// TIA Portal V17 program export: 0 tag tables, 0 data types, 5 data blocks, 5 code blocks (in call order from the OBs), 4 instance data blocks

DATA_BLOCK "DB_HMI"   // DB1
{ S7_Optimized_Access := 'TRUE' }
VERSION : 0.1
// stored: AutoNumber true, DBAccessibleFromOPCUA true, IsOnlyStoredInLoadMemory false, IsRetainMemResEnabled false, IsWriteProtectedInAS false, MemoryReserve 100
   VAR
      Cmd_Marcha : Bool;   // Boton MARCHA de la HMI (momentaneo)
      Cmd_Paro : Bool;   // Boton PARO de la HMI (momentaneo)
      Cmd_Reset : Bool;   // Boton RESET de la HMI (momentaneo)
      Sel_Estilo : Int := 1;   // 1 Banderas, 2 Moore, 3 Mealy
      Estado : Int;   // Estado del estilo seleccionado: 0 Reposo, 10 Marcha, 90 Falla
      Motor_En_Marcha : Bool;   // Copia de KM1_Motor para la HMI
      Falla_Termico : Bool;   // Termico disparado
      Pantalla : Int;   // Pantalla activa en la HMI (1 Principal, 2 Diagnostico, 3 Estilos)
   END_VAR
BEGIN
END_DATA_BLOCK

DATA_BLOCK "DB_Mando"
{ S7_Optimized_Access := 'TRUE' }
VERSION : 0.1
NON_RETAIN
"FB_Mando_Motor"

BEGIN

END_DATA_BLOCK

DATA_BLOCK "DB_Motor_Banderas"
{ S7_Optimized_Access := 'TRUE' }
VERSION : 0.1
NON_RETAIN
"FB_Motor_Banderas"

BEGIN

END_DATA_BLOCK

DATA_BLOCK "DB_Motor_Mealy"
{ S7_Optimized_Access := 'TRUE' }
VERSION : 0.1
NON_RETAIN
"FB_Motor_Mealy"

BEGIN

END_DATA_BLOCK

DATA_BLOCK "DB_Motor_Moore"
{ S7_Optimized_Access := 'TRUE' }
VERSION : 0.1
NON_RETAIN
"FB_Motor_Moore"

BEGIN

END_DATA_BLOCK

ORGANIZATION_BLOCK "Main"   // OB1, LAD, ProgramCycle
TITLE = "Main Program Sweep (Cycle)" / Programa principal - Arranque y paro v2
{ S7_Optimized_Access := 'TRUE' }
VERSION : 0.1
// OB1 director: una red por función. Los 3 estilos corren a la vez; el selector de la HMI decide cuál maneja KM1 y los pilotos.
// stored: AutoNumber true, IsIECCheckEnabled false, SetENOAutomatically false
   VAR_INPUT
      Initial_Call : Bool;   // Initial call of this OB
      Remanence : Bool;   // =True, if remanent data are available
   END_VAR
BEGIN

REGION Network 1: MANDO: pulsadores + HMI
   // Une entradas físicas y botones de la HMI.
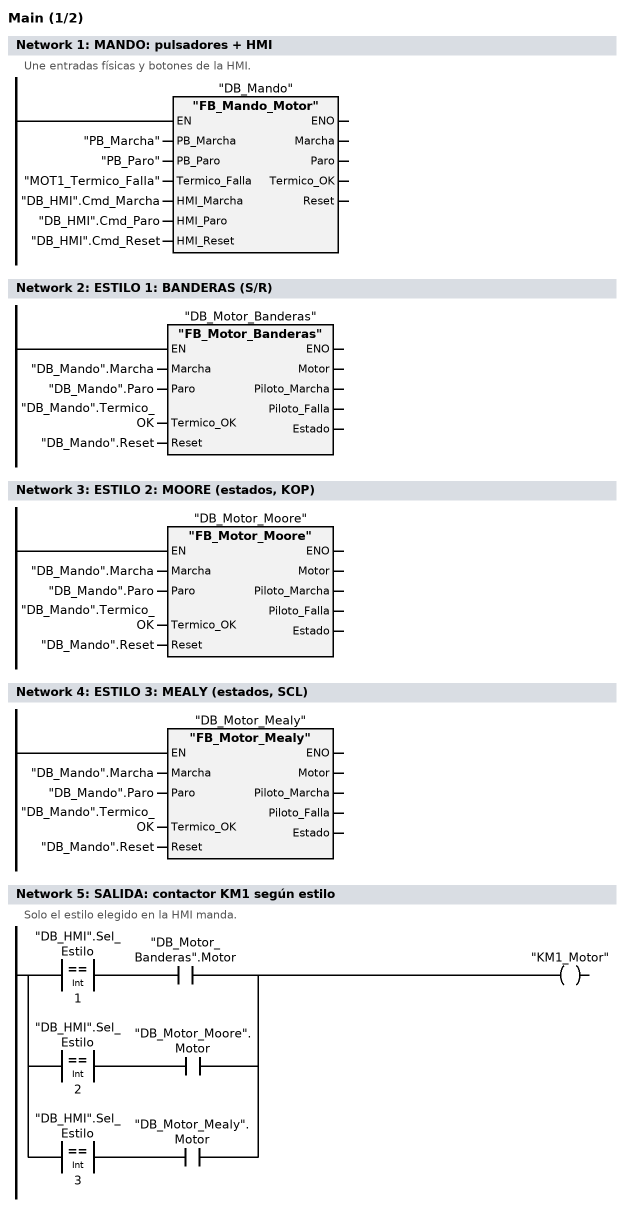
   RUNG wire#powerrail
      "DB_Mando"(PB_Marcha := "PB_Marcha", PB_Paro := "PB_Paro", Termico_Falla := "MOT1_Termico_Falla", HMI_Marcha := "DB_HMI".Cmd_Marcha, HMI_Paro := "DB_HMI".Cmd_Paro, HMI_Reset := "DB_HMI".Cmd_Reset, Marcha =>, Paro =>, Termico_OK =>, Reset =>)
   END_RUNG
   // the same network as SCL:
   "DB_Mando"(PB_Marcha := "PB_Marcha",   // "FB_Mando_Motor"
              PB_Paro := "PB_Paro",
              Termico_Falla := "MOT1_Termico_Falla",
              HMI_Marcha := "DB_HMI".Cmd_Marcha,
              HMI_Paro := "DB_HMI".Cmd_Paro,
              HMI_Reset := "DB_HMI".Cmd_Reset);
END_REGION

REGION Network 2: ESTILO 1: BANDERAS (S/R)
   RUNG wire#powerrail
      "DB_Motor_Banderas"(Marcha := "DB_Mando".Marcha, Paro := "DB_Mando".Paro, Termico_OK := "DB_Mando".Termico_OK, Reset := "DB_Mando".Reset, Motor =>, Piloto_Marcha =>, Piloto_Falla =>, Estado =>)
   END_RUNG
   // the same network as SCL:
   "DB_Motor_Banderas"(Marcha := "DB_Mando".Marcha,   // "FB_Motor_Banderas"
                       Paro := "DB_Mando".Paro,
                       Termico_OK := "DB_Mando".Termico_OK,
                       Reset := "DB_Mando".Reset);
END_REGION

REGION Network 3: ESTILO 2: MOORE (estados, KOP)
   RUNG wire#powerrail
      "DB_Motor_Moore"(Marcha := "DB_Mando".Marcha, Paro := "DB_Mando".Paro, Termico_OK := "DB_Mando".Termico_OK, Reset := "DB_Mando".Reset, Motor =>, Piloto_Marcha =>, Piloto_Falla =>, Estado =>)
   END_RUNG
   // the same network as SCL:
   "DB_Motor_Moore"(Marcha := "DB_Mando".Marcha,   // "FB_Motor_Moore"
                    Paro := "DB_Mando".Paro,
                    Termico_OK := "DB_Mando".Termico_OK,
                    Reset := "DB_Mando".Reset);
END_REGION

REGION Network 4: ESTILO 3: MEALY (estados, SCL)
   RUNG wire#powerrail
      "DB_Motor_Mealy"(Marcha := "DB_Mando".Marcha, Paro := "DB_Mando".Paro, Termico_OK := "DB_Mando".Termico_OK, Reset := "DB_Mando".Reset, Motor =>, Piloto_Marcha =>, Piloto_Falla =>, Estado =>)
   END_RUNG
   // the same network as SCL:
   "DB_Motor_Mealy"(Marcha := "DB_Mando".Marcha,   // "FB_Motor_Mealy"
                    Paro := "DB_Mando".Paro,
                    Termico_OK := "DB_Mando".Termico_OK,
                    Reset := "DB_Mando".Reset);
END_REGION

REGION Network 5: SALIDA: contactor KM1 según estilo
   // Solo el estilo elegido en la HMI manda.
   RUNG wire#powerrail
      { S7_Templates := "SrcType := Int" } EQ_Contact(in1 := "DB_HMI".Sel_Estilo, in2 := 1)
      Contact( "DB_Motor_Banderas".Motor )
      wire#w1
      Coil( "KM1_Motor" )
   END_RUNG
   RUNG wire#powerrail
      { S7_Templates := "SrcType := Int" } EQ_Contact(in1 := "DB_HMI".Sel_Estilo, in2 := 2)
      Contact( "DB_Motor_Moore".Motor )
   END_RUNG wire#w1
   RUNG wire#powerrail
      { S7_Templates := "SrcType := Int" } EQ_Contact(in1 := "DB_HMI".Sel_Estilo, in2 := 3)
      Contact( "DB_Motor_Mealy".Motor )
   END_RUNG wire#w1
   // the same network as SCL:
   "KM1_Motor" := (("DB_HMI".Sel_Estilo = 1) AND "DB_Motor_Banderas".Motor) OR (("DB_HMI".Sel_Estilo = 2) AND "DB_Motor_Moore".Motor) OR (("DB_HMI".Sel_Estilo = 3) AND "DB_Motor_Mealy".Motor);
END_REGION

REGION Network 6: SALIDA: piloto de marcha
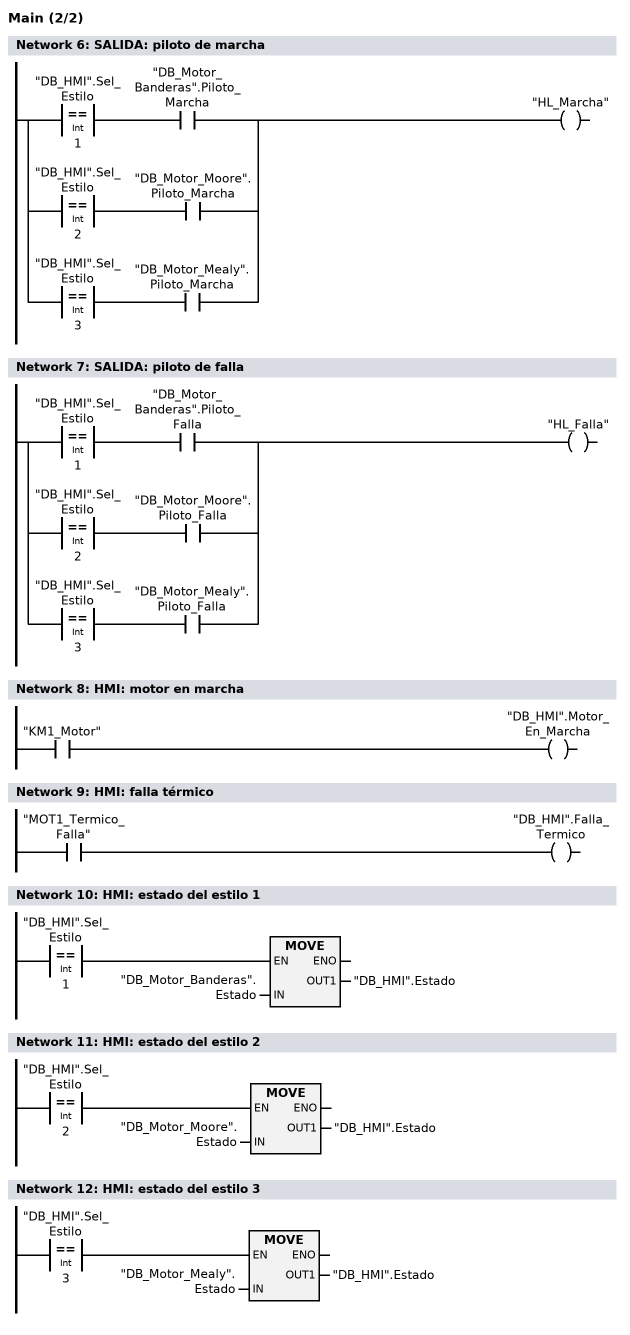
   RUNG wire#powerrail
      { S7_Templates := "SrcType := Int" } EQ_Contact(in1 := "DB_HMI".Sel_Estilo, in2 := 1)
      Contact( "DB_Motor_Banderas".Piloto_Marcha )
      wire#w1
      Coil( "HL_Marcha" )
   END_RUNG
   RUNG wire#powerrail
      { S7_Templates := "SrcType := Int" } EQ_Contact(in1 := "DB_HMI".Sel_Estilo, in2 := 2)
      Contact( "DB_Motor_Moore".Piloto_Marcha )
   END_RUNG wire#w1
   RUNG wire#powerrail
      { S7_Templates := "SrcType := Int" } EQ_Contact(in1 := "DB_HMI".Sel_Estilo, in2 := 3)
      Contact( "DB_Motor_Mealy".Piloto_Marcha )
   END_RUNG wire#w1
   // the same network as SCL:
   "HL_Marcha" := (("DB_HMI".Sel_Estilo = 1) AND "DB_Motor_Banderas".Piloto_Marcha) OR (("DB_HMI".Sel_Estilo = 2) AND "DB_Motor_Moore".Piloto_Marcha) OR (("DB_HMI".Sel_Estilo = 3) AND "DB_Motor_Mealy".Piloto_Marcha);
END_REGION

REGION Network 7: SALIDA: piloto de falla
   RUNG wire#powerrail
      { S7_Templates := "SrcType := Int" } EQ_Contact(in1 := "DB_HMI".Sel_Estilo, in2 := 1)
      Contact( "DB_Motor_Banderas".Piloto_Falla )
      wire#w1
      Coil( "HL_Falla" )
   END_RUNG
   RUNG wire#powerrail
      { S7_Templates := "SrcType := Int" } EQ_Contact(in1 := "DB_HMI".Sel_Estilo, in2 := 2)
      Contact( "DB_Motor_Moore".Piloto_Falla )
   END_RUNG wire#w1
   RUNG wire#powerrail
      { S7_Templates := "SrcType := Int" } EQ_Contact(in1 := "DB_HMI".Sel_Estilo, in2 := 3)
      Contact( "DB_Motor_Mealy".Piloto_Falla )
   END_RUNG wire#w1
   // the same network as SCL:
   "HL_Falla" := (("DB_HMI".Sel_Estilo = 1) AND "DB_Motor_Banderas".Piloto_Falla) OR (("DB_HMI".Sel_Estilo = 2) AND "DB_Motor_Moore".Piloto_Falla) OR (("DB_HMI".Sel_Estilo = 3) AND "DB_Motor_Mealy".Piloto_Falla);
END_REGION

REGION Network 8: HMI: motor en marcha
   RUNG wire#powerrail
      Contact( "KM1_Motor" )
      Coil( "DB_HMI".Motor_En_Marcha )
   END_RUNG
   // the same network as SCL:
   "DB_HMI".Motor_En_Marcha := "KM1_Motor";
END_REGION

REGION Network 9: HMI: falla térmico
   RUNG wire#powerrail
      Contact( "MOT1_Termico_Falla" )
      Coil( "DB_HMI".Falla_Termico )
   END_RUNG
   // the same network as SCL:
   "DB_HMI".Falla_Termico := "MOT1_Termico_Falla";
END_REGION

REGION Network 10: HMI: estado del estilo 1
   RUNG wire#powerrail
      { S7_Templates := "SrcType := Int" } EQ_Contact(in1 := "DB_HMI".Sel_Estilo, in2 := 1)
      { S7_GenerateENO := "TRUE" } Move(in := "DB_Motor_Banderas".Estado, out1 => "DB_HMI".Estado)
   END_RUNG
   // the same network as SCL:
   IF "DB_HMI".Sel_Estilo = 1 THEN "DB_HMI".Estado := "DB_Motor_Banderas".Estado; END_IF;
END_REGION

REGION Network 11: HMI: estado del estilo 2
   RUNG wire#powerrail
      { S7_Templates := "SrcType := Int" } EQ_Contact(in1 := "DB_HMI".Sel_Estilo, in2 := 2)
      { S7_GenerateENO := "TRUE" } Move(in := "DB_Motor_Moore".Estado, out1 => "DB_HMI".Estado)
   END_RUNG
   // the same network as SCL:
   IF "DB_HMI".Sel_Estilo = 2 THEN "DB_HMI".Estado := "DB_Motor_Moore".Estado; END_IF;
END_REGION

REGION Network 12: HMI: estado del estilo 3
   RUNG wire#powerrail
      { S7_Templates := "SrcType := Int" } EQ_Contact(in1 := "DB_HMI".Sel_Estilo, in2 := 3)
      { S7_GenerateENO := "TRUE" } Move(in := "DB_Motor_Mealy".Estado, out1 => "DB_HMI".Estado)
   END_RUNG
   // the same network as SCL:
   IF "DB_HMI".Sel_Estilo = 3 THEN "DB_HMI".Estado := "DB_Motor_Mealy".Estado; END_IF;
END_REGION
END_ORGANIZATION_BLOCK

FUNCTION_BLOCK "FB_Mando_Motor"   // FB1, LAD
TITLE = Mando del motor: pulsadores + HMI
{ S7_Optimized_Access := 'TRUE' }
VERSION : 0.1
// Une pulsadores físicos y botones HMI. Reset = botón RESET de la HMI o mantener MARCHA 3 s.
// stored: AutoNumber true, IsIECCheckEnabled false, IsRetainMemResEnabled false, MemoryReserve 100, SetENOAutomatically false, UDAEnableTagReadback false
   VAR_INPUT
      PB_Marcha : Bool;   // Pulsador MARCHA (NA)
      PB_Paro : Bool;   // Pulsador PARO: 1 = pulsado
      Termico_Falla : Bool;   // Relé térmico: 1 = disparado
      HMI_Marcha : Bool;
      HMI_Paro : Bool;
      HMI_Reset : Bool;
   END_VAR
   VAR_OUTPUT
      Marcha : Bool;
      Paro : Bool;
      Termico_OK : Bool;
      Reset : Bool;
   END_VAR
   VAR
      T_Reset : TON_TIME;   // Tiempo de MARCHA mantenida
      Reset_Mantenido : Bool;   // MARCHA mantenida 3 s
   END_VAR
BEGIN

REGION Network 1: Marcha
   // Pulsador físico o botón de la HMI.
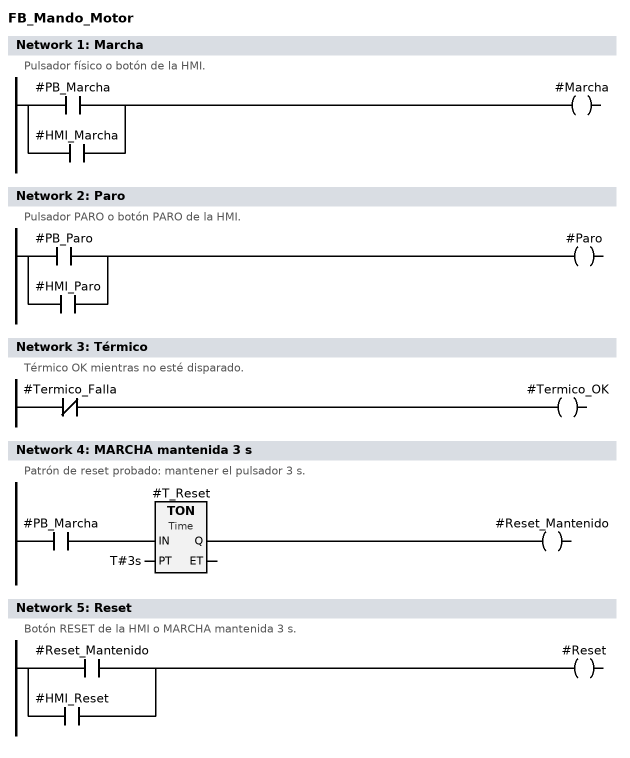
   RUNG wire#powerrail
      Contact( #PB_Marcha )
      wire#w1
      Coil( #Marcha )
   END_RUNG
   RUNG wire#powerrail
      Contact( #HMI_Marcha )
   END_RUNG wire#w1
   // the same network as SCL:
   #Marcha := #PB_Marcha OR #HMI_Marcha;
END_REGION

REGION Network 2: Paro
   // Pulsador PARO o botón PARO de la HMI.
   RUNG wire#powerrail
      Contact( #PB_Paro )
      wire#w1
      Coil( #Paro )
   END_RUNG
   RUNG wire#powerrail
      Contact( #HMI_Paro )
   END_RUNG wire#w1
   // the same network as SCL:
   #Paro := #PB_Paro OR #HMI_Paro;
END_REGION

REGION Network 3: Térmico
   // Térmico OK mientras no esté disparado.
   RUNG wire#powerrail
      I_Contact( #Termico_Falla )
      Coil( #Termico_OK )
   END_RUNG
   // the same network as SCL:
   #Termico_OK := NOT #Termico_Falla;
END_REGION

REGION Network 4: MARCHA mantenida 3 s
   // Patrón de reset probado: mantener el pulsador 3 s.
   RUNG wire#powerrail
      Contact( #PB_Marcha )
      { S7_Templates := "time_type := Time" } #T_Reset.TON(pt := T#3s, et =>)
      Coil( #Reset_Mantenido )
   END_RUNG
   // the same network as SCL:
   #T_Reset(IN := #PB_Marcha, PT := T#3s);   // TON
   #Reset_Mantenido := #T_Reset.Q;
END_REGION

REGION Network 5: Reset
   // Botón RESET de la HMI o MARCHA mantenida 3 s.
   RUNG wire#powerrail
      Contact( #Reset_Mantenido )
      wire#w1
      Coil( #Reset )
   END_RUNG
   RUNG wire#powerrail
      Contact( #HMI_Reset )
   END_RUNG wire#w1
   // the same network as SCL:
   #Reset := #Reset_Mantenido OR #HMI_Reset;
END_REGION
END_FUNCTION_BLOCK

FUNCTION_BLOCK "FB_Motor_Banderas"   // FB3, LAD
TITLE = Arranque y paro por BANDERAS (S/R)
{ S7_Optimized_Access := 'TRUE' }
VERSION : 0.1
// Estilo clásico: bandera de marcha con SET/RESET (paro dominante). Sin térmico se para; al recuperarse el térmico se puede volver a arrancar sin RESET.
// stored: AutoNumber true, IsIECCheckEnabled false, IsRetainMemResEnabled false, MemoryReserve 100, SetENOAutomatically false, UDAEnableTagReadback false
   VAR_INPUT
      Marcha : Bool;   // Orden de marcha (pulsador o HMI)
      Paro : Bool;   // Orden de paro: 1 = parar
      Termico_OK : Bool;   // 1 = relé térmico sin falla
      Reset : Bool;   // Reset de falla
   END_VAR
   VAR_OUTPUT
      Motor : Bool;   // Orden al contactor
      Piloto_Marcha : Bool;   // Piloto verde
      Piloto_Falla : Bool;   // Piloto rojo
      Estado : Int;   // 0 Reposo, 10 Marcha, 90 Falla
   END_VAR
   VAR
      B_Marcha : Bool;   // Bandera: motor en marcha
      B_Falla : Bool;   // Bandera: falla térmico
   END_VAR
BEGIN

REGION Network 1: SET bandera de marcha
   // Marcha sin paro y con térmico OK.
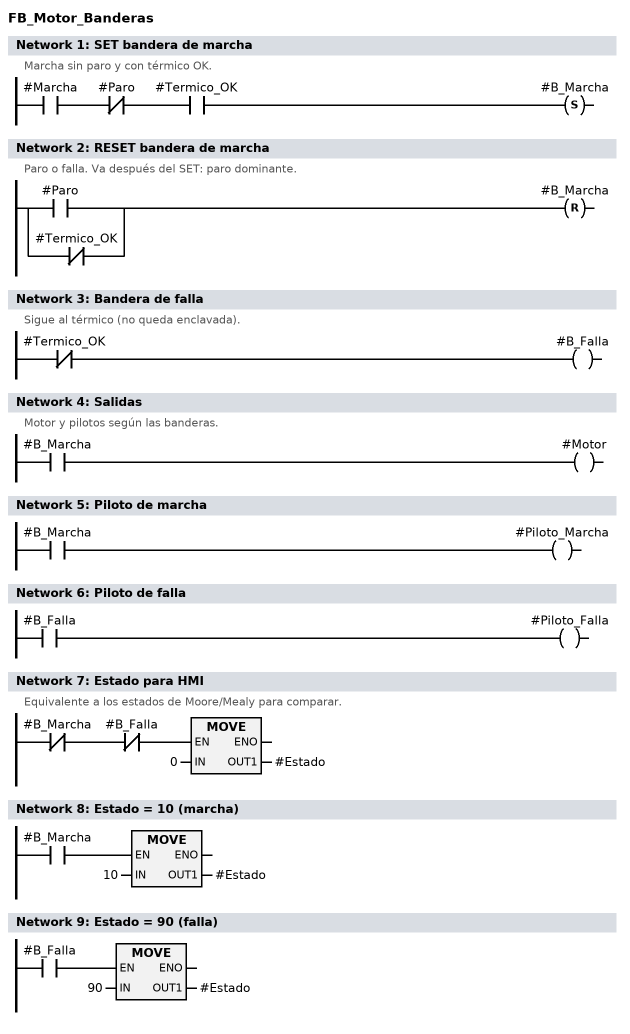
   RUNG wire#powerrail
      Contact( #Marcha )
      I_Contact( #Paro )
      Contact( #Termico_OK )
      S_Coil( #B_Marcha )
   END_RUNG
   // the same network as SCL:
   IF #Marcha AND NOT #Paro AND #Termico_OK THEN #B_Marcha := TRUE; END_IF;
END_REGION

REGION Network 2: RESET bandera de marcha
   // Paro o falla. Va después del SET: paro dominante.
   RUNG wire#powerrail
      Contact( #Paro )
      wire#w1
      R_Coil( #B_Marcha )
   END_RUNG
   RUNG wire#powerrail
      I_Contact( #Termico_OK )
   END_RUNG wire#w1
   // the same network as SCL:
   IF #Paro OR NOT #Termico_OK THEN #B_Marcha := FALSE; END_IF;
END_REGION

REGION Network 3: Bandera de falla
   // Sigue al térmico (no queda enclavada).
   RUNG wire#powerrail
      I_Contact( #Termico_OK )
      Coil( #B_Falla )
   END_RUNG
   // the same network as SCL:
   #B_Falla := NOT #Termico_OK;
END_REGION

REGION Network 4: Salidas
   // Motor y pilotos según las banderas.
   RUNG wire#powerrail
      Contact( #B_Marcha )
      Coil( #Motor )
   END_RUNG
   // the same network as SCL:
   #Motor := #B_Marcha;
END_REGION

REGION Network 5: Piloto de marcha
   RUNG wire#powerrail
      Contact( #B_Marcha )
      Coil( #Piloto_Marcha )
   END_RUNG
   // the same network as SCL:
   #Piloto_Marcha := #B_Marcha;
END_REGION

REGION Network 6: Piloto de falla
   RUNG wire#powerrail
      Contact( #B_Falla )
      Coil( #Piloto_Falla )
   END_RUNG
   // the same network as SCL:
   #Piloto_Falla := #B_Falla;
END_REGION

REGION Network 7: Estado para HMI
   // Equivalente a los estados de Moore/Mealy para comparar.
   RUNG wire#powerrail
      I_Contact( #B_Marcha )
      I_Contact( #B_Falla )
      { S7_GenerateENO := "TRUE" } Move(in := 0, out1 => #Estado)
   END_RUNG
   // the same network as SCL:
   IF NOT #B_Marcha AND NOT #B_Falla THEN #Estado := 0; END_IF;
END_REGION

REGION Network 8: Estado = 10 (marcha)
   RUNG wire#powerrail
      Contact( #B_Marcha )
      { S7_GenerateENO := "TRUE" } Move(in := 10, out1 => #Estado)
   END_RUNG
   // the same network as SCL:
   IF #B_Marcha THEN #Estado := 10; END_IF;
END_REGION

REGION Network 9: Estado = 90 (falla)
   RUNG wire#powerrail
      Contact( #B_Falla )
      { S7_GenerateENO := "TRUE" } Move(in := 90, out1 => #Estado)
   END_RUNG
   // the same network as SCL:
   IF #B_Falla THEN #Estado := 90; END_IF;
END_REGION
END_FUNCTION_BLOCK

FUNCTION_BLOCK "FB_Motor_Moore"   // FB5, LAD
TITLE = Arranque y paro: máquina de estados MOORE
{ S7_Optimized_Access := 'TRUE' }
VERSION : 0.1
// Moore: las salidas dependen solo del estado. Generado por TIA_MCP_V17 (crear_maquina_estados).
// stored: AutoNumber true, IsIECCheckEnabled false, IsRetainMemResEnabled false, MemoryReserve 100, SetENOAutomatically false, UDAEnableTagReadback false
   VAR_INPUT
      Marcha : Bool;   // Orden de marcha (pulsador o HMI)
      Paro : Bool;   // Orden de paro: 1 = parar
      Termico_OK : Bool;   // 1 = relé térmico sin falla
      Reset : Bool;   // Reset de falla
   END_VAR
   VAR_OUTPUT
      Motor : Bool;   // Orden al contactor
      Piloto_Marcha : Bool;   // Piloto verde
      Piloto_Falla : Bool;   // Piloto rojo
      Estado : Int;   // Estado actual
   END_VAR
   VAR
      Estado_Actual : Int := 0;   // Estado de la máquina
   END_VAR
   VAR_TEMP
      Estado_Previo : Int;   // Estado al inicio del ciclo
   END_VAR
BEGIN

REGION Network 1: Foto del estado al inicio del ciclo
   // Las transiciones se evalúan sobre esta copia: un solo salto por ciclo.
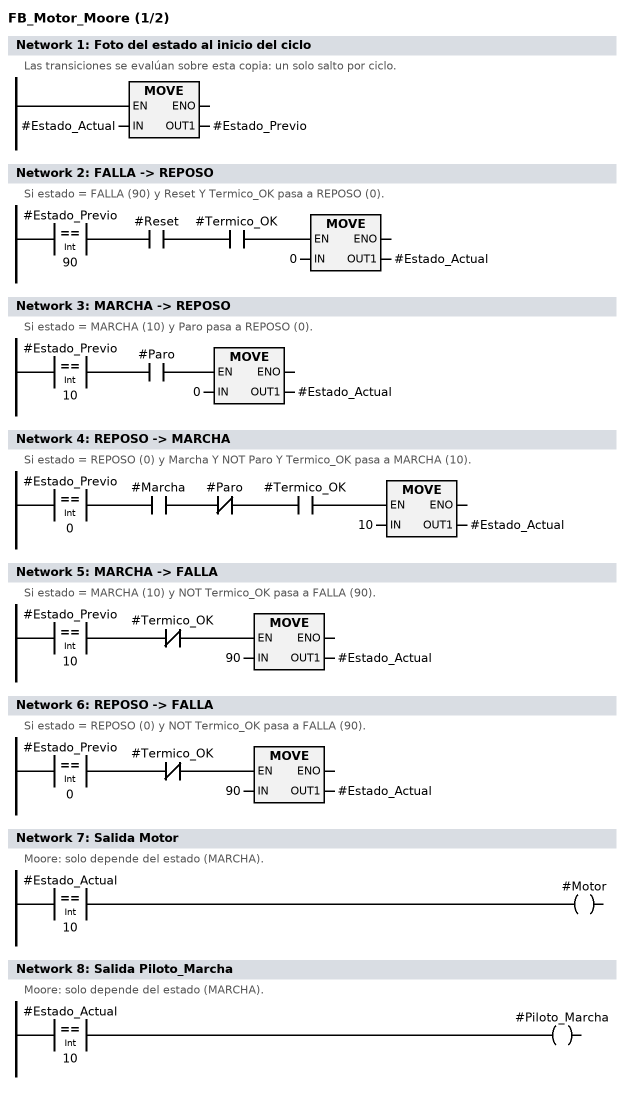
   RUNG wire#powerrail
      { S7_GenerateENO := "TRUE" } Move(in := #Estado_Actual, out1 => #Estado_Previo)
   END_RUNG
   // the same network as SCL:
   #Estado_Previo := #Estado_Actual;
END_REGION

REGION Network 2: FALLA -> REPOSO
   // Si estado = FALLA (90) y Reset Y Termico_OK pasa a REPOSO (0).
   RUNG wire#powerrail
      { S7_Templates := "SrcType := Int" } EQ_Contact(in1 := #Estado_Previo, in2 := 90)
      Contact( #Reset )
      Contact( #Termico_OK )
      { S7_GenerateENO := "TRUE" } Move(in := 0, out1 => #Estado_Actual)
   END_RUNG
   // the same network as SCL:
   IF (#Estado_Previo = 90) AND #Reset AND #Termico_OK THEN #Estado_Actual := 0; END_IF;
END_REGION

REGION Network 3: MARCHA -> REPOSO
   // Si estado = MARCHA (10) y Paro pasa a REPOSO (0).
   RUNG wire#powerrail
      { S7_Templates := "SrcType := Int" } EQ_Contact(in1 := #Estado_Previo, in2 := 10)
      Contact( #Paro )
      { S7_GenerateENO := "TRUE" } Move(in := 0, out1 => #Estado_Actual)
   END_RUNG
   // the same network as SCL:
   IF (#Estado_Previo = 10) AND #Paro THEN #Estado_Actual := 0; END_IF;
END_REGION

REGION Network 4: REPOSO -> MARCHA
   // Si estado = REPOSO (0) y Marcha Y NOT Paro Y Termico_OK pasa a MARCHA (10).
   RUNG wire#powerrail
      { S7_Templates := "SrcType := Int" } EQ_Contact(in1 := #Estado_Previo, in2 := 0)
      Contact( #Marcha )
      I_Contact( #Paro )
      Contact( #Termico_OK )
      { S7_GenerateENO := "TRUE" } Move(in := 10, out1 => #Estado_Actual)
   END_RUNG
   // the same network as SCL:
   IF (#Estado_Previo = 0) AND #Marcha AND NOT #Paro AND #Termico_OK THEN #Estado_Actual := 10; END_IF;
END_REGION

REGION Network 5: MARCHA -> FALLA
   // Si estado = MARCHA (10) y NOT Termico_OK pasa a FALLA (90).
   RUNG wire#powerrail
      { S7_Templates := "SrcType := Int" } EQ_Contact(in1 := #Estado_Previo, in2 := 10)
      I_Contact( #Termico_OK )
      { S7_GenerateENO := "TRUE" } Move(in := 90, out1 => #Estado_Actual)
   END_RUNG
   // the same network as SCL:
   IF (#Estado_Previo = 10) AND NOT #Termico_OK THEN #Estado_Actual := 90; END_IF;
END_REGION

REGION Network 6: REPOSO -> FALLA
   // Si estado = REPOSO (0) y NOT Termico_OK pasa a FALLA (90).
   RUNG wire#powerrail
      { S7_Templates := "SrcType := Int" } EQ_Contact(in1 := #Estado_Previo, in2 := 0)
      I_Contact( #Termico_OK )
      { S7_GenerateENO := "TRUE" } Move(in := 90, out1 => #Estado_Actual)
   END_RUNG
   // the same network as SCL:
   IF (#Estado_Previo = 0) AND NOT #Termico_OK THEN #Estado_Actual := 90; END_IF;
END_REGION

REGION Network 7: Salida Motor
   // Moore: solo depende del estado (MARCHA).
   RUNG wire#powerrail
      { S7_Templates := "SrcType := Int" } EQ_Contact(in1 := #Estado_Actual, in2 := 10)
      Coil( #Motor )
   END_RUNG
   // the same network as SCL:
   #Motor := #Estado_Actual = 10;
END_REGION

REGION Network 8: Salida Piloto_Marcha
   // Moore: solo depende del estado (MARCHA).
   RUNG wire#powerrail
      { S7_Templates := "SrcType := Int" } EQ_Contact(in1 := #Estado_Actual, in2 := 10)
      Coil( #Piloto_Marcha )
   END_RUNG
   // the same network as SCL:
   #Piloto_Marcha := #Estado_Actual = 10;
END_REGION

REGION Network 9: Salida Piloto_Falla
   // Moore: solo depende del estado (FALLA).
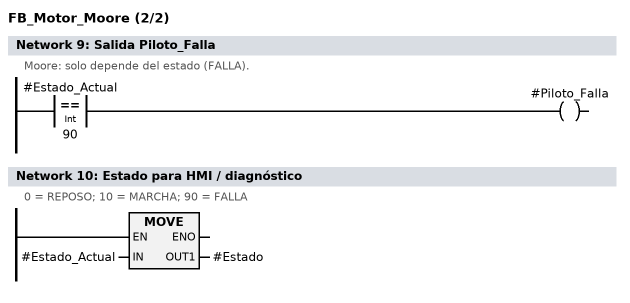
   RUNG wire#powerrail
      { S7_Templates := "SrcType := Int" } EQ_Contact(in1 := #Estado_Actual, in2 := 90)
      Coil( #Piloto_Falla )
   END_RUNG
   // the same network as SCL:
   #Piloto_Falla := #Estado_Actual = 90;
END_REGION

REGION Network 10: Estado para HMI / diagnóstico
   // 0 = REPOSO; 10 = MARCHA; 90 = FALLA
   RUNG wire#powerrail
      { S7_GenerateENO := "TRUE" } Move(in := #Estado_Actual, out1 => #Estado)
   END_RUNG
   // the same network as SCL:
   #Estado := #Estado_Actual;
END_REGION
END_FUNCTION_BLOCK

FUNCTION_BLOCK "FB_Motor_Mealy"   // FB4, SCL
TITLE = Arranque y paro: maquina de estados MEALY
{ S7_Optimized_Access := 'TRUE' }
VERSION : 0.1
// stored: AutoNumber true, IsIECCheckEnabled false, IsRetainMemResEnabled false, MemoryReserve 100, SetENOAutomatically false, UDAEnableTagReadback false
   VAR_INPUT
      Marcha : Bool;   // Orden de marcha (pulsador o HMI)
      Paro : Bool;   // Orden de paro: 1 = parar
      Termico_OK : Bool;   // 1 = rele termico sin falla
      Reset : Bool;   // Reset de falla
   END_VAR
   VAR_OUTPUT
      Motor : Bool;   // Orden al contactor
      Piloto_Marcha : Bool;   // Piloto verde
      Piloto_Falla : Bool;   // Piloto rojo
      Estado : Int;   // Estado actual (HMI)
   END_VAR
   VAR
      Estado_Actual : Int := 0;   // Estado de la maquina
   END_VAR
   VAR_TEMP
      Estado_Previo : Int;   // Estado al inicio del ciclo
   END_VAR
BEGIN
       // Mealy: las salidas dependen del estado y de las entradas (reaccion en el mismo ciclo). Generado por TIA_MCP_V17 (crear_maquina_estados).
       // Estados: 0 = REPOSO, 10 = MARCHA, 90 = FALLA

       // --- Salidas (estado actual + entradas) ---
       #Motor := (#Estado_Actual = 10 AND NOT #Paro AND #Termico_OK);
       #Piloto_Marcha := #Estado_Actual = 10;
       #Piloto_Falla := #Estado_Actual = 90;

       // --- Transiciones (sobre la foto del estado: un salto por ciclo) ---
       #Estado_Previo := #Estado_Actual;
       CASE #Estado_Previo OF
           0: // REPOSO
               IF NOT #Termico_OK THEN
                   #Estado_Actual := 90;   // -> FALLA
               ELSIF #Marcha AND NOT #Paro AND #Termico_OK THEN
                   #Estado_Actual := 10;   // -> MARCHA
               END_IF;
           10: // MARCHA
               IF NOT #Termico_OK THEN
                   #Estado_Actual := 90;   // -> FALLA
               ELSIF #Paro THEN
                   #Estado_Actual := 0;   // -> REPOSO
               END_IF;
           90: // FALLA
               IF #Reset AND #Termico_OK THEN
                   #Estado_Actual := 0;   // -> REPOSO
               END_IF;
           ELSE  // estado desconocido: volver al inicial
               #Estado_Actual := 0;
       END_CASE;

       #Estado := #Estado_Actual;
END_FUNCTION_BLOCK

DATA_BLOCK "DB_Mando"   // DB2
VERSION : 0.1
// stored: AutoNumber true, DBAccessibleFromOPCUA true, InstanceOfName FB_Mando_Motor, InstanceOfType FB
"FB_Mando_Motor"
BEGIN
END_DATA_BLOCK

DATA_BLOCK "DB_Motor_Banderas"   // DB3
VERSION : 0.1
// stored: AutoNumber true, DBAccessibleFromOPCUA true, InstanceOfName FB_Motor_Banderas, InstanceOfType FB
"FB_Motor_Banderas"
BEGIN
END_DATA_BLOCK

DATA_BLOCK "DB_Motor_Mealy"   // DB5
VERSION : 0.1
// stored: AutoNumber true, DBAccessibleFromOPCUA true, InstanceOfName FB_Motor_Mealy, InstanceOfType FB
"FB_Motor_Mealy"
BEGIN
END_DATA_BLOCK

DATA_BLOCK "DB_Motor_Moore"   // DB4
VERSION : 0.1
// stored: AutoNumber true, DBAccessibleFromOPCUA true, InstanceOfName FB_Motor_Moore, InstanceOfType FB
"FB_Motor_Moore"
BEGIN
END_DATA_BLOCK
